{attribute 'no_explicit_call' := 'Direct call not allowed for type FB_TurCtl'}
{attribute 'call_after_init'}
FUNCTION_BLOCK FB_TurCtl EXTENDS FB_AcsiBATypeENUMERATED
VAR
	_eValue: E_TurCtl;
	_eConfig: E_TurCtl;
	{attribute 'hide'}
	ipInit: I_AcsiCommonAttributeClass := THIS^.AddDAValue(eP:=E_AcsiP.Actual, in:=_eValue).AddDAValue(eP:=E_AcsiP.Config, in:=_eConfig).AddDAType(in:=THIS^.T(in:=E_AcsiBasicType.INT8));
END_VAR

PROPERTY eConfig : E_TurCtl
GET
eConfig:= _eConfig;
END_GET
END_PROPERTY

PROPERTY eValue : E_TurCtl
GET
eValue:= _eValue;
OnGetVPropEvt();
END_GET
SET
_bChanged:= _eValue <> eValue;
_eValue:= eValue;
OnSetVPropEvt(bChanged := _bChanged);
END_SET
END_PROPERTY

END_FUNCTION_BLOCK

(* stored: Version 1.1.0.1
   POU FB_TurCtl: Id {8ffe8840-0404-4177-b001-afde18597c30}, SpecialFunc None
   Property eConfig: Id {f81479d6-e285-4fde-91d8-d6dbec33e6aa}
   Get Get: Id {e3e7eaca-3967-4353-b394-8d8cd6941113}
   Property eValue: Id {5ec521aa-5004-454d-8016-4e51195c5f90}
   Get Get: Id {052ef588-bd1a-45b9-a9ec-c2c196ed1297}
   Set Set: Id {308b74e6-1d61-4b24-b0fc-a695d26c63c1} *)
